ABB RobotStudio station: NeuralTest.rsstn

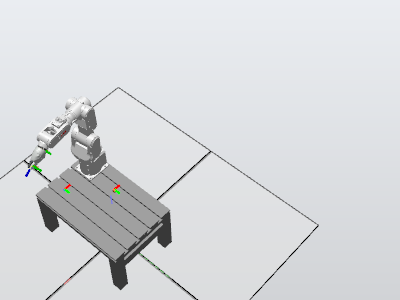
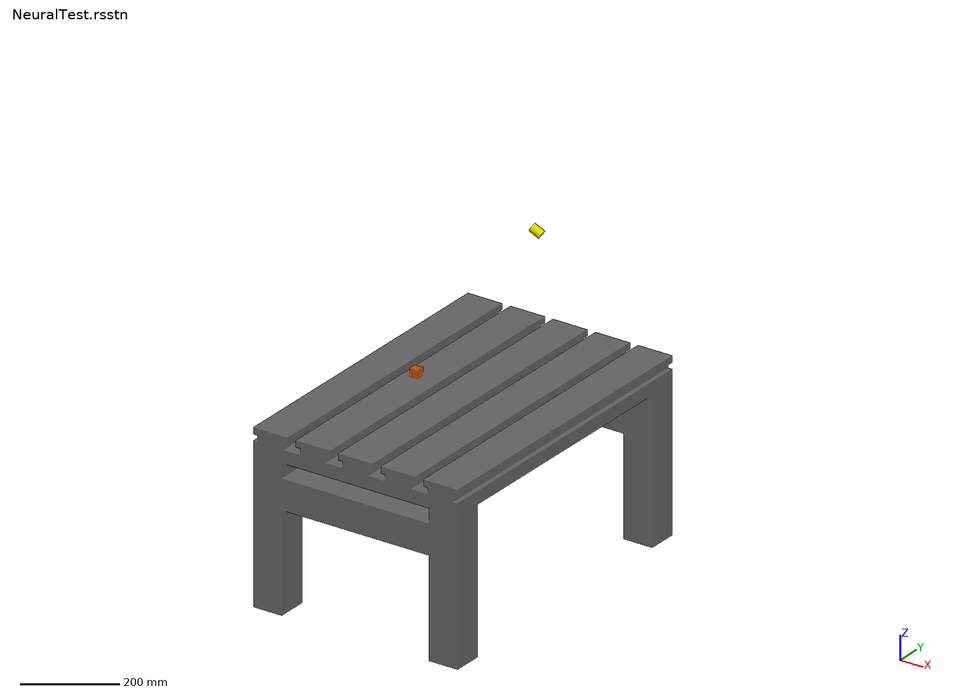
[picture v1: parts stored in the station drawn from their meshes, with robot base, taught points and paths (robot models come from the ABB library and are not in the file)]
Station Station (saved by RobotStudio 26.3.11844.1)
Layout (positions relative to the parent item):
  - Table_small [part] at (-218.8, -434.83, 0) mm, size 500 x 750 x 400 mm
  - IRB1100_4_58_BTM_01 [mechanism, from %ABB.RobotStudio.Models.IRB1100%\IRB1100_4_58_BTM_01.rslib] at (-111.22, -315.19, 404.46) mm; joint values [0.1256, 0, 0, 0, 0.5236, 0] (rad or m)
  - Smart_Gripper_Servo_Fingers [mechanism, from %ABB.RobotStudio.Models.SmartGripper%\ABB_Smart_Gripper_Servo_Fingers.rslib] at (241.41, -270.66, 989.46) mm, rotated rx 180 ry 60 rz -172.8 deg; joint values [0.025] (rad or m)
  - LineSensor [smart component, from Components\LineSensor.rslib] at (339.53, -258.28, 932.36) mm, rotated rx 180 ry 60 rz -172.8 deg
      properties: Start=[0 0 0]; End=[0 0 0.025]; Length=0.025; Radius=0.010000000000000002; Tag=(none); SenseMultiple=false; SensedPart=(none); SensedPoint=[0 0 0]
    - _sensorPart_ [part], size 20 x 20 x 25 mm
  - Attacher [smart component, from Components\Attacher.rslib]
      properties: Parent=(none); Flange=0; Child=(none); Mount=false; Offset=[0 0 0]; Orientation=[0 0 0]
  - Detacher [smart component, from Components\Detacher.rslib]
      properties: Child=(none); KeepPosition=true
  - box [part] at (-112.8, -89.83, 380.84) mm, size 20 x 20 x 20 mm
Attachment: Smart_Gripper_Servo_Fingers is attached to IRB1100_4_58_BTM_01 / Link6
Attachment: LineSensor is attached to Smart_Gripper_Servo_Fingers / HandBase
Station logic (signal -> signal, property => property):
  LineSensor.SensedPart => Attacher.Child
  Attacher.Child => Detacher.Child
Targets, tools, work objects and paths stored in the station, written as RAPID:
! task (no controller)
MODULE Module1
  CONST robtarget Target_center:=[[-82.8,-59.827,420.838],[0,0,1,0],[0,0,0,0],[9E+09,9E+09,9E+09,9E+09,9E+09,9E+09]];
  CONST robtarget Target_side:=[[134.607257778,-306.182858465,423.952983979],[0,0,1,0],[0,0,0,0],[9E+09,9E+09,9E+09,9E+09,9E+09,9E+09]];
ENDMODULE

! task (no controller)
MODULE CalibData
  PERS tooldata Servo:=[TRUE,[[0,0,114.2],[1,0,0,0]],[0.215,[8.7,12.3,49.2],[1,0,0,0],0.00021,0.00024,0.00009]];
ENDMODULE

! task (no controller)
MODULE Module1
  CONST jointtarget Home:=[[0,0,0,0,90,0],[9E+09,9E+09,9E+09,9E+09,9E+09,9E+09]];
ENDMODULE

